% RSLogix 500 project Traffic Light Cycle2_BAK018.RSS, saved by version 8.30.00.16 %
PROJECT "PLCLAB"    % processor: Bul.1763 MicroLogix 1100 Series B %

PROGRAM FILES
  LAD 2 "MAIN"  5 rungs
  LAD 3 "DIGITAL IO"  6 rungs
  LAD 4 "ANALOG IO"  1 rungs
  LAD 5 "ALARMS"  1 rungs
  LAD 6 "CONTROLS"  6 rungs

DATA FILES
  O0 OUTPUT  5 elements
  I1 INPUT  7 elements
  S2 STATUS  66 elements
  B3 BINARY  1 elements
  T4 TIMER  4 elements
  C5 COUNTER  1 elements
  R6 CONTROL  1 elements
  N7 INTEGER  1 elements
  F8 FLOAT  1 elements

LADDER 2 "MAIN"
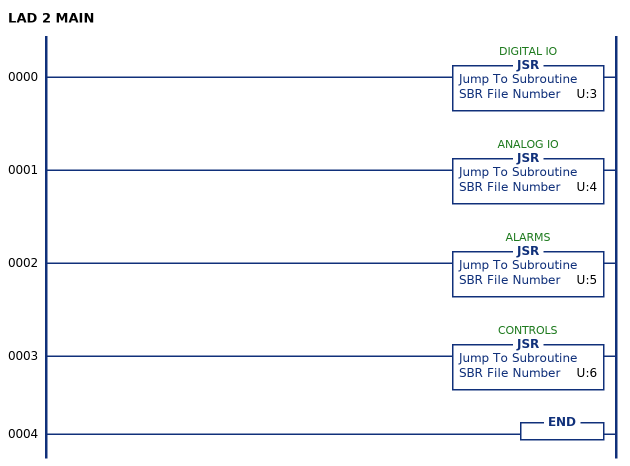
% Rung: 0 %
SOR JSR U:3 EOR
%   U:3  "DIGITAL IO" %
% Rung: 1 %
SOR JSR U:4 EOR
%   U:4  "ANALOG IO" %
% Rung: 2 %
SOR JSR U:5 EOR
%   U:5  "ALARMS" %
% Rung: 3 %
SOR JSR U:6 EOR
%   U:6  "CONTROLS" %
% Rung: 4 %
SOR END EOR

LADDER 3 "DIGITAL IO"
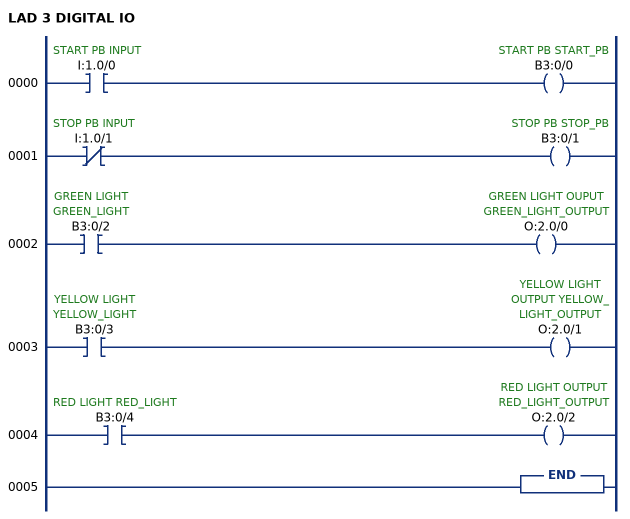
% Rung: 0 %
SOR XIC I:1.0/0 OTE B3:0/0 EOR
%   I:1.0/0  "START PB INPUT" %
%   B3:0/0  START_PB  "START PB" %
% Rung: 1 %
SOR XIO I:1.0/1 OTE B3:0/1 EOR
%   I:1.0/1  "STOP PB INPUT" %
%   B3:0/1  STOP_PB  "STOP PB" %
% Rung: 2 %
SOR XIC B3:0/2 OTE O:2.0/0 EOR
%   B3:0/2  GREEN_LIGHT  "GREEN LIGHT" %
%   O:2.0/0  GREEN_LIGHT_OUTPUT  "GREEN LIGHT OUPUT" %
% Rung: 3 %
SOR XIC B3:0/3 OTE O:2.0/1 EOR
%   B3:0/3  YELLOW_LIGHT  "YELLOW LIGHT" %
%   O:2.0/1  YELLOW_LIGHT_OUTPUT  "YELLOW LIGHT OUTPUT" %
% Rung: 4 %
SOR XIC B3:0/4 OTE O:2.0/2 EOR
%   B3:0/4  RED_LIGHT  "RED LIGHT" %
%   O:2.0/2  RED_LIGHT_OUTPUT  "RED LIGHT OUTPUT" %
% Rung: 5 %
SOR END EOR

LADDER 6 "CONTROLS"
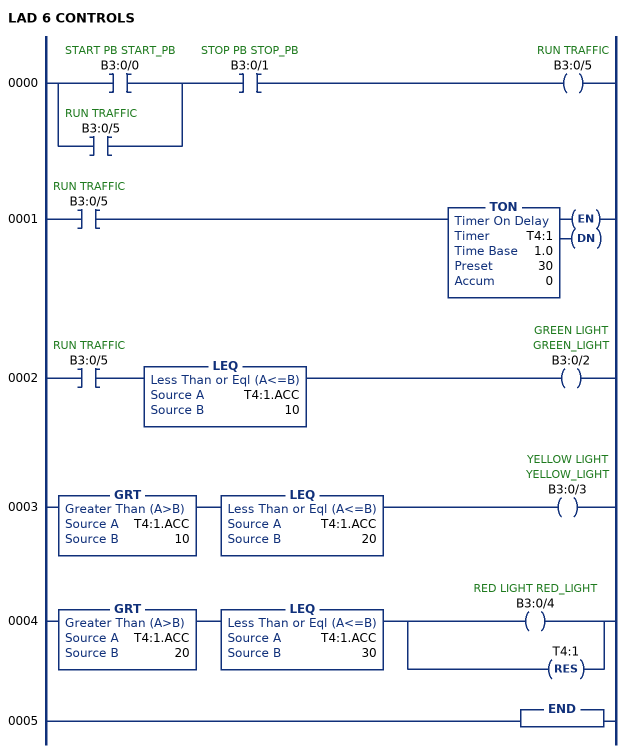
% Rung: 0 %
SOR BST XIC B3:0/0 NXB XIC B3:0/5 BND XIC B3:0/1 OTE B3:0/5 EOR
%   B3:0/0  START_PB  "START PB" %
%   B3:0/5  "RUN TRAFFIC" %
%   B3:0/1  STOP_PB  "STOP PB" %
% Rung: 1 %
SOR XIC B3:0/5 TON T4:1 1.0 30 0 EOR
%   B3:0/5  "RUN TRAFFIC" %
% Rung: 2 %
SOR XIC B3:0/5 LEQ T4:1.ACC 10 OTE B3:0/2 EOR
%   B3:0/5  "RUN TRAFFIC" %
%   B3:0/2  GREEN_LIGHT  "GREEN LIGHT" %
% Rung: 3 %
SOR GRT T4:1.ACC 10 LEQ T4:1.ACC 20 OTE B3:0/3 EOR
%   B3:0/3  YELLOW_LIGHT  "YELLOW LIGHT" %
% Rung: 4 %
SOR GRT T4:1.ACC 20 LEQ T4:1.ACC 30 BST OTE B3:0/4 NXB RES T4:1 BND EOR
%   B3:0/4  RED_LIGHT  "RED LIGHT" %
% Rung: 5 %
SOR END EOR

OTHER DOCUMENTED ADDRESSES
  I:0.0/2  "GREEN INPUT LIGHT"
  I:1.0/2  "GREEN INPUT LIGHT"
  I:1.0/3  "YELLOW INPUT LIGHT"
  I:1.0/4  "RED INPUT LIGHT"
  LEQ  
  T4:0  "GREEN LIGHT TIMER"

DATA TABLE (non-zero values as saved)
DATA T4
% .PRE .ACC %
% T4:0 % 10 0
% T4:1 % 30 0
% T4:2 % 10 0
% T4:3 % 10 0
